Fanuc KAREL source: kt00238.KL

-- PROVISIONAL review KL for V770-1; original PC SHA256 2b2ec4e50843a88b8e6b43673b868271a9aa68af4614b7865d75050ccb2d2727
-- Incomplete behavior may be omitted. Consult companion uncertainty JSON. Do not deploy.
PROGRAM KT00238
%NOLOCKGROUP
VAR
  I1 : INTEGER
  OUT : INTEGER
-- UNRESOLVED_DECL Y2 type=002018
BEGIN
  -- UNRESOLVED_PC offsets 5-16; opcodes 2E,23
  -- UNRESOLVED_PC offsets 21-35; opcodes 2E,22,9D,33,B2
  -- UNRESOLVED_PC offsets 40-62; opcodes 21,22,9D,33,B1,47,23
  -- UNRESOLVED_PC offsets 67-71; opcodes 7F
END KT00238
